FUNCTION FUN_Write_Line_To_History : BOOL
VAR_INPUT
END_VAR
VAR
	i: INT;
END_VAR

	FOR i:=C_Max_Buffer_Act_list TO 2 BY -1 DO
		Buffer_Act_History[i]:=Buffer_Act_History[i-1];
	END_FOR
	Buffer_Act_History[1]:=Buffer_Act_Message[1];

END_FUNCTION

(* stored: Version 1.1.0.1, ProductVersion 3.1.4024.15
   POU FUN_Write_Line_To_History: Id {2bbab7bb-9998-4057-b64e-98d4fa1a7ed8}, SpecialFunc None *)
